Fanuc KAREL source: ka00068.KL

-- PROVISIONAL review KL for V770-1; original PC SHA256 82c2c88e1822143b7bbc786d875a0ac4337c20a949c79e703ba9abaaa3e71f91
-- Incomplete behavior may be omitted. Consult companion uncertainty JSON. Do not deploy.
PROGRAM KA00068
%NOLOCKGROUP
-- UNRESOLVED_DECL SRC type=000102
-- UNRESOLVED_DECL DST type=000199
BEGIN
  -- UNRESOLVED_PC offsets 5-20; opcodes 2E,22,32,35
  -- UNRESOLVED_PC offsets 25-45; opcodes 49,7E,4A
  -- UNRESOLVED_PC offsets 50-54; opcodes 7F
END KA00068
